RoboDK station: ronan.rdk

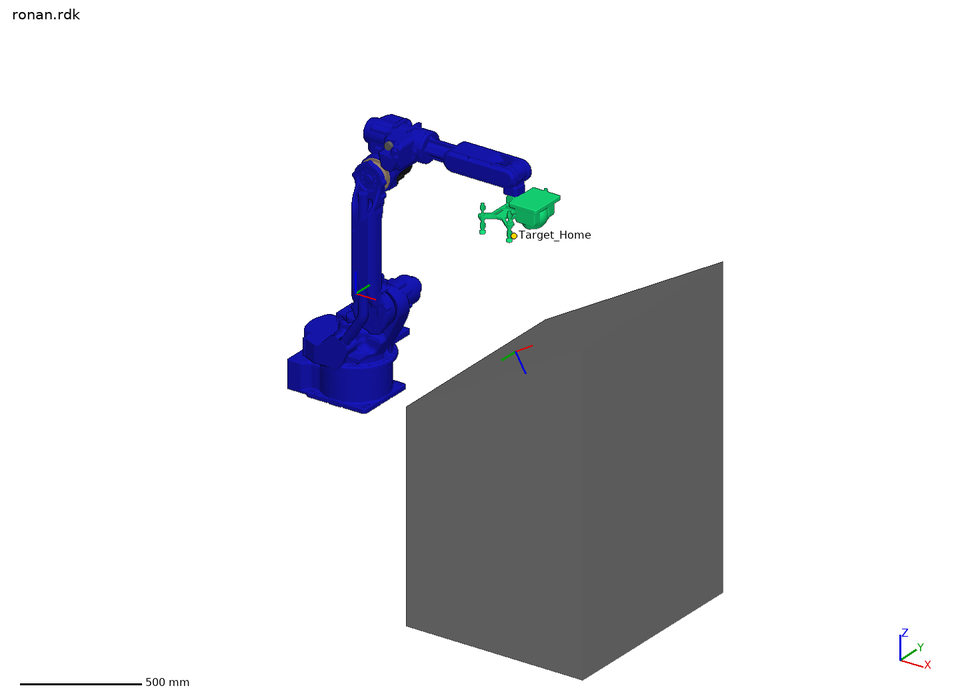
[picture v0: the station drawn from its stored meshes, robots at their saved joint values, targets as dots, program paths as lines]
Station Robodk (2) (saved by RoboDK 6.1.1). Poses are relative to the parent item; angles as X-Y-Z fixed-axis rotations.
  - frame Motoman MH6 Base at (0, 0, 450) mm
    - robot Motoman MH6: 6 axes, payload 6 kg, reach 1422 mm, repeatability 0.08 mm, weight 130 kg
        modified DH rows (alpha deg, a mm, theta deg, d mm): 0, 0, 0, 450; -90, 152, -90, 0; 0, 614, 0, 0; -90, 155, 0, 640; 90, 0, 90, 0; -90, 0, 0, 95
        base shift (0, 0, -450) mm
        joint limits [-170, -90, -175, -180, -45, -360] to [170, 155, 250, 180, 225, 360]; home [0, 0, 0, 0, 0, 0]; saved at [0, 0, 0, 0, 0, 0]
      - tool Ventosas, TCP at (0, 0, 190) mm, size 250 x 290 x 148 mm
    - frame Frame_from_Target1 at (823.2, -34.49, -21.13) mm, rotated rx -180 ry -30 rz 0 deg
      - target Target_Home (Cartesian target) at (225.55, -34.49, -453.06) mm, rotated rx 0 ry -30 rz 0 deg; joints [0, 0, 0, 0, 0, 0] of Motoman MH6
  - object CAJA2 at (1600, 500, 300) mm, rotated rx 180 ry 0 rz 0 deg, size 886.4 x 1000 x 1511.7 mm, geometry from CAJA2.stp
  - Python program RosPolar (listed below)
  - Python program Prog2 (listed below)

--- Python program RosPolar ---
from robodk.robolink import *    # API para comunicarte con RoboDK
from robodk.robomath import *    # Funciones matemáticas
import math

#------------------------------------------------
# 1) Conexión a RoboDK e inicialización
#------------------------------------------------
RDK = Robolink()

# Elegir un robot (si hay varios, aparece un popup)
robot = RDK.ItemUserPick("Selecciona un robot", ITEM_TYPE_ROBOT)
if not robot.Valid():
    raise Exception("No se ha seleccionado un robot válido.")

# Conectar al robot físico
#if not robot.Connect():
#    raise Exception("No se pudo conectar al robot. Verifica que esté en modo remoto y que la configuración sea correcta.")

# Confirmar conexión
#if not robot.ConnectedState():
#    raise Exception("El robot no está conectado correctamente. Revisa la conexión.")

print("Robot conectado correctamente.")

#------------------------------------------------
# 2) Cargar el Frame (ya existente) donde quieres dibujar
#    Ajusta el nombre si tu Frame se llama diferente
#------------------------------------------------
frame_name = "Frame_from_Target1"
frame = RDK.Item(frame_name, ITEM_TYPE_FRAME)
home = "Target_Home"
homeFM = RDK.Item(home, ITEM_TYPE_TARGET)
if not frame.Valid():
    raise Exception(f'No se encontró el Frame "{frame_name}" en la estación.')

# Asignamos este frame al robot
robot.setPoseFrame(frame)
# Usamos la herramienta activa
robot.setPoseTool(robot.PoseTool())

# Ajustes de velocidad y blending
robot.setSpeed(300)   # mm/s - Ajusta según necesites
robot.setRounding(5)  # blending (radio de curvatura)

#------------------------------------------------
# 3) Parámetros de la figura (rosa polar)
#------------------------------------------------
num_points = 720       # Cuántos puntos muestreamos (mayor = más suave)
A = 150               # Amplitud (300 mm = radio máximo)
k = 5                  # Parámetro de la rosa (pétalos). Si es impar, habrá k pétalos; si es par, 2k
z_surface = 0          # Z=0 en el plano del frame
z_safe = 50            # Altura segura para aproximarse y salir

#------------------------------------------------
# 4) Movimiento al centro en altura segura
#------------------------------------------------

robot.MoveJ(homeFM)
# El centro de la rosa (r=0) corresponde a x=0, y=0
robot.MoveJ(transl(0, 0, z_surface - z_safe))

# Bajamos a la "superficie" (Z=0)
robot.MoveL(transl(0, 0, z_surface))

#------------------------------------------------
# 5) Dibujar la rosa polar
#    r = A * sin(k*theta)
#    x = r*cos(theta), y = r*sin(theta)
#------------------------------------------------
# Recorremos theta de 0 a 2*pi (una vuelta completa)
full_turn = 24*math.pi

for i in range(num_points+1):
    # Fracción entre 0 y 1
    t = i / num_points
    # Ángulo actual
    theta = full_turn * t

    # Calculamos r
    r = (
    math.exp(math.sin(theta))
    - 2 * math.cos(4 * theta)
    + math.sin((2 * theta - math.pi) / 24) ** 5
    + 0.5 * math.sin(8 * theta) * math.cos(theta / 8) ** 2
   )
    # Convertimos a coordenadas Cartesianas X, Y
    x = r * math.cos(theta)
    y = r * math.sin(theta)

    # Movemos linealmente (MoveL) en el plano del Frame
    robot.MoveL(transl(x, y, z_surface))

# Al terminar, subimos de nuevo para no chocar
robot.MoveL(transl(x, y, z_surface - z_safe))
robot.MoveJ(homeFM)
print(f"¡Figura (rosa polar) completada en el frame '{frame_name}'!")

--- Python program Prog2 ---
from robodk.robolink import *
from robodk.robomath import *
import math
from matplotlib.textpath import TextPath
from matplotlib.font_manager import FontProperties
from matplotlib.textpath import TextToPath


#------------------------------------------------
# 1) Connexion à RoboDK
#------------------------------------------------
RDK = Robolink()

robot = RDK.ItemUserPick("Selecciona un robot", ITEM_TYPE_ROBOT)
if not robot.Valid():
    raise Exception("No se ha seleccionado un robot válido.")


# Conectar al robot físico
#if not robot.Connect():
#    raise Exception("No se pudo conectar al robot. Verifica que esté en modo remoto y que la configuración sea correcta.")

# Confirmar conexión
#if not robot.ConnectedState():
#    raise Exception("El robot no está conectado correctamente. Revisa la conexión.")


#------------------------------------------------
# 2) Frame y target home
#------------------------------------------------
frame_name = "Frame_from_Target1"
frame = RDK.Item(frame_name, ITEM_TYPE_FRAME)
homeFM = RDK.Item("Target_Home", ITEM_TYPE_TARGET)
if not frame.Valid():
    raise Exception(f'No se encontró el Frame "{frame_name}" en la estación.')
if not homeFM.Valid():
    raise Exception('No se encontró "Target_Home".')

robot.setPoseFrame(frame)
robot.setPoseTool(robot.PoseTool())
robot.setSpeed(300)     # mm/s
robot.setRounding(1)    # blending pequeño (segmentos muy cortos)

#------------------------------------------------
# 3) Parámetros de la figura
#------------------------------------------------
num_points = 50          # puntos de la curva (3000-5000 va bien)
A = 150                    # radio máximo deseado en mm
z_surface = 0
z_safe = 50                # si tu eje Z del frame apunta hacia arriba, usa +z_safe

# Orientación de la herramienta respecto al frame.
# Si el robot no llega o la herramienta apunta al revés, prueba: rotx(math.pi)
orient = eye(4)

def pose_xyz(x, y, z):
    return transl(x, y, z) * orient

#------------------------------------------------
# 4) Calcular la curva (θ de 0 a 24π)
#------------------------------------------------
def r_func(theta):
    return (
        math.exp(math.sin(theta))
        - 2 * math.cos(4 * theta)
        + math.sin((2 * theta - math.pi) / 24) ** 5
        + 0.5 * math.sin(8 * theta) * math.cos(theta / 8) ** 2
    )

full_turn = 24 * math.pi
thetas = [full_turn * i / num_points for i in range(num_points + 1)]
radios = [r_func(t) for t in thetas]

# Escalamos para que el radio máximo sea A mm
scale = A / max(abs(r) for r in radios)

puntos = [(scale * r * math.cos(t), scale * r * math.sin(t))
          for r, t in zip(radios, thetas)]

#------------------------------------------------
# 5) Movimiento
#------------------------------------------------
robot.MoveJ(homeFM)

# Ir encima del primer punto en altura segura, luego bajar
x0, y0 = puntos[0]
robot.MoveJ(pose_xyz(x0, y0, z_surface - z_safe))
robot.MoveL(pose_xyz(x0, y0, z_surface))

fp = FontProperties(family="sans", style="italic")
path1, codes = TextToPath().get_text_path(fp, "Alejandro")
path2, codes = TextToPath().get_text_path(fp, "Nirvana")
path3, codes = TextToPath().get_text_path(fp, "Ronan")

for punto in path1:
    x,y=punto
    robot.MoveL(pose_xyz(y+400,x-path1[-1][0], z_surface))
for punto in path2:
    x,y=punto
    robot.MoveL(pose_xyz(y+300,x-path2[-1][0], z_surface))
for punto in path3:
    x,y=punto
    robot.MoveL(pose_xyz(y+200,x-path3[-1][0], z_surface))


# Dibujar
for (x, y) in puntos:
    robot.MoveL(pose_xyz(x, y, z_surface))



# Subir y volver a home
xf, yf = puntos[-1]
robot.MoveL(pose_xyz(xf, yf, z_surface - z_safe))
robot.MoveJ(homeFM)

print(f"¡Figura completada en el frame '{frame_name}'! (escala = {scale:.2f} mm/unidad)")
